FUNCTION_BLOCK FB_Delayed
VAR_INPUT
    enable : BOOL;
    delay : TIME := T#1s;
END_VAR
VAR_OUTPUT
    ready : BOOL;
    elapsed : TIME;
END_VAR
VAR
    delayTimer : TON;
END_VAR

delayTimer(IN := enable, PT := delay, Q => ready, ET => elapsed);

END_FUNCTION_BLOCK

(* stored: Version 1.1.0.1 *)
